(* IEC 61131-3 sources: bottling-plant/pous/function-blocks, 13 files *)

(* ---- BangBangControl.st ---- *)
FUNCTION_BLOCK BangBangControl
  VAR
    Hysteresis : HYSTERESIS;
  END_VAR
  VAR_INPUT
    Setpoint : REAL;
    Tolerance : REAL;
  END_VAR
  VAR_OUTPUT
    Readback : REAL;
    ShouldActuate : DINT;
  END_VAR

Hysteresis( XIN1 := Setpoint, XIN2 := Readback, EPS := Tolerance);
ShouldActuate := Hysteresis.Q;

END_FUNCTION_BLOCK

(* ---- FB_11_MixingTank.st ---- *)
FUNCTION_BLOCK FB_11_MixingTank
  VAR
    TempControl : BANGBANGCONTROL;
    LevelControl : BANGBANGCONTROL;
    RequestTempControl : BOOL;
    RequestLevelControl : BOOL;
    LatchingFault : LATCHINGFAULT;
    OpenInlet : BOOL;
    HeaterOn : BOOL;
  END_VAR
  VAR_INPUT
  END_VAR
  VAR_OUTPUT
    LevelReadback : REAL;
  END_VAR

TempControl(Tolerance := 1);
LevelControl(Tolerance := 0.2);

LatchingFault(Active := RequestTempControl AND RequestLevelControl);

HeaterOn := RequestTempControl AND TempControl.ShouldActuate AND NOT LatchingFault.LatchedOutput;
OpenInlet := RequestLevelControl AND LevelControl.ShouldActuate AND NOT LatchingFault.LatchedOutput;
LevelReadback := LevelControl.Readback;

END_FUNCTION_BLOCK

(* ---- FB_12_TransferPump.st ---- *)
FUNCTION_BLOCK FB_12_TransferPump
  VAR
    RequestMixDrain : BOOL;
    MixOutletOpen : BOOL;
  END_VAR
  VAR CONSTANT
  END_VAR
  VAR_INPUT
    MixLevelReadback : REAL;
  END_VAR
  VAR_TEMP
  END_VAR
  VAR_OUTPUT
    BufferLevelReadback : REAL;
    LatchingFault : LATCHINGFAULT;
  END_VAR

MixOutletOpen := RequestMixDrain AND MixLevelReadback > 1 AND NOT LatchingFault.LatchedOutput;

END_FUNCTION_BLOCK

(* ---- FB_1_Process.st ---- *)
FUNCTION_BLOCK FB_1_Process
  VAR
    MixingTank : FB_11_MIXINGTANK;
    TransferPump : FB_12_TRANSFERPUMP;
  END_VAR
  VAR_OUTPUT
    BufferLevel : REAL;
  END_VAR

MixingTank();
TransferPump(MixLevelReadback := MixingTank.LevelReadback);
BufferLevel := TransferPump.BufferLevelReadback;

END_FUNCTION_BLOCK

(* ---- FB_2_Packaging.st ---- *)
FUNCTION_BLOCK FB_2_Packaging
  VAR
    Filler : FB_2_PACKAGING_FILLER;
    Conveyor : FB_2_PACKAGING_CONVEYOR;
  END_VAR

Filler();
Conveyor();

END_FUNCTION_BLOCK

(* ---- FB_2_Packaging_Conveyor.st ---- *)
FUNCTION_BLOCK FB_2_Packaging_Conveyor
  VAR
    LoadBottle : BOOL;
    BottleLoaded : BOOL;
    CompressedAirReadback : BOOL;
    CoolingLoopReadback : BOOL;
  END_VAR
  VAR_INPUT
  END_VAR

END_FUNCTION_BLOCK

(* ---- FB_2_Packaging_Filler.st ---- *)
FUNCTION_BLOCK FB_2_Packaging_Filler
  VAR
    FlowRateSetpoint_mm3_s : REAL;
    FlowRateReadback_mm3_s : REAL;
    FillVolume_mm3 : REAL;
    CompressedAirReadback : REAL;
    CoolingLoopReadback : REAL;
  END_VAR
  VAR_OUTPUT
  END_VAR

if FillVolume_mm3 > 100 then
    BottleFull := TRUE;
end_if
OverFillFault(Active := FillVolume_mm3 > 120);

END_FUNCTION_BLOCK

(* ---- FB_3_Motion.st ---- *)
FUNCTION_BLOCK FB_3_Motion
  VAR
    Capper : FB_3_MOTION_CAPPER;
    CasePacker : FB_3_MOTION_CASEPACKER;
  END_VAR

Capper();
CasePacker();

END_FUNCTION_BLOCK

(* ---- FB_3_Motion_Capper.st ---- *)
FUNCTION_BLOCK FB_3_Motion_Capper
  VAR
    ApplyTorque : REAL;
    AngularVelocityFeedback : REAL;
    AngleFeedback : REAL;
    ResistTorqueFeedback : REAL;
    CompressedAirReadback : REAL;
    CoolingLoopReadback : REAL;
  END_VAR

END_FUNCTION_BLOCK

(* ---- FB_3_Motion_CasePacker.st ---- *)
FUNCTION_BLOCK FB_3_Motion_CasePacker
  VAR
    InitiatePack : BOOL;
    PackState : BOOL;
    BottleCount : DINT;
    CaseCount : DINT;
  END_VAR

END_FUNCTION_BLOCK

(* ---- FB_4_Utilities.st ---- *)
FUNCTION_BLOCK FB_4_Utilities
  VAR
    CompressedAir : FB_4_UTILITIES_FACILITYUTILITY;
    CoolingLoop : FB_4_UTILITIES_FACILITYUTILITY;
  END_VAR

CompressedAir();
CoolingLoop();

END_FUNCTION_BLOCK

(* ---- FB_4_Utilities_FacilityUtility.st ---- *)
FUNCTION_BLOCK FB_4_Utilities_FacilityUtility
  VAR
    GenerationSetpoint : REAL;
    GenerationReadback : REAL;
    TargetReadback : REAL;
  END_VAR
  VAR_INPUT
  END_VAR

END_FUNCTION_BLOCK

(* ---- LatchingFault.st ---- *)
FUNCTION_BLOCK LatchingFault
  VAR
  END_VAR
  VAR_INPUT
    Active : BOOL := FALSE;
    Reset : BOOL := FALSE;
  END_VAR
  VAR_OUTPUT
    LatchedOutput : BOOL := FALSE;
  END_VAR

LatchedOutput := Active OR (LatchedOutput AND NOT Reset);

END_FUNCTION_BLOCK
